Fanuc KAREL source: KX00013.KL

PROGRAM KX00013
%NOLOCKGROUP
VAR
  I: INTEGER
  J: INTEGER
  B: BOOLEAN
  F: FILE
  S: STRING[80]
  P: XYZWPR
BEGIN
  RESUME
END KX00013
